(* IEC 61131-3 sources: SortJet_MasterSPS_Aufbau.fbsproj/07_Auftragsverwaltung/SystemCheck.prg.st^, 7 files *)

(* ---- Auftraege_Shuttle.meth.st ---- *)
(* METADATA
{
	"v3Meta": {
		"objectGuid": "9ff2d478-3fef-409c-b42e-3dce6a33e4ba"
	}
}
*)
METHOD PRIVATE Auftraege_Shuttle : BOOL
VAR_INPUT
  wpAutomatikkreis : WORD;
END_VAR

//-------------------------------------------------------------------------------------------------
// SYSTEMCHECK - AUTOMATIKKREIS 1
//-------------------------------------------------------------------------------------------------

Auftraege_Shuttle := FALSE;

FOR wlIndex := cERSTES_SHUTTLE TO cLETZTES_SHUTTLE DO
  IF wpAutomatikkreis = starrShuttleBasisParameter[wlIndex].stMKs.eaAutomatikkreis[1] THEN
    IF starrShuttleBasisParameter[wlIndex].stMKs.eStationsTyp = eInputshuttle THEN//101,102
      CASE starrShuttleBasisParameter[wlIndex].pAuftrag[cWAND_1].wTransferstationsNr1 OF

        cERSTE_STATION..cLETZTE_STATION:
          starrShuttleBasisParameter[wlIndex].pAuftrag[cWAND_1].stAuftragsOptionen.eGlastransport := eGlastransport_AufEinlaufVorab;
          starrShuttleBasisParameter[wlIndex].pAuftrag[cWAND_1].stAuftragsOptionen.eKippen_SollPosition := eKippen_Position_90Grad;
          Auftraege_Shuttle := TRUE;

        cERSTES_TRANSFERSHUTTLE..cLETZTES_TRANSFERSHUTTLE,
        cSPEICHER_1..cSPEICHER_2:
          starrShuttleBasisParameter[wlIndex].pAuftrag[cWAND_1].stAuftragsOptionen.eGlastransport := eGlastransport_AufAuslauf;
          starrShuttleBasisParameter[wlIndex].pAuftrag[cWAND_1].stAuftragsOptionen.eKippen_SollPosition := eKippen_Position_90Grad;//1.5
          Auftraege_Shuttle := TRUE;

        cERSTE_FAECHERWAGENSTATIONS_NR..cLETZTE_FAECHERWAGENSTATIONS_NR:
          starrShuttleBasisParameter[wlIndex].pAuftrag[cWAND_1].stAuftragsOptionen.eGlastransport := eGlastransport_AufAuslauf;
          starrShuttleBasisParameter[wlIndex].pAuftrag[cWAND_1].stAuftragsOptionen.eKippen_SollPosition := eKippen_Position_90Grad;
          Auftraege_Shuttle := TRUE;

        ELSE
          starrShuttleBasisParameter[wlIndex].pAuftrag[cWAND_1].stAuftragsOptionen.eGlastransport := eGlastransport_AufAuslauf;
          starrShuttleBasisParameter[wlIndex].pAuftrag[cWAND_1].stAuftragsOptionen.eKippen_SollPosition := eKippen_Position_90Grad;
          Auftraege_Shuttle := TRUE;

      END_CASE

    ELSIF starrShuttleBasisParameter[wlIndex].stMKs.eStationsTyp = eOutputshuttle THEN//103,104
      CASE starrShuttleBasisParameter[wlIndex].pAuftrag[cWAND_1].wTransferstationsNr1 OF

        cERSTES_TRANSFERSHUTTLE..cLETZTES_TRANSFERSHUTTLE,
        cSPEICHER_1:
          starrShuttleBasisParameter[wlIndex].pAuftrag[cWAND_1].stAuftragsOptionen.eGlastransport := eGlastransport_AufEinlaufVorab;
          starrShuttleBasisParameter[wlIndex].pAuftrag[cWAND_1].stAuftragsOptionen.eKippen_SollPosition := eKippen_Position_90Grad;//1.5
          Auftraege_Shuttle := TRUE;

        cERSTE_STATION..cLETZTE_STATION:
          starrShuttleBasisParameter[wlIndex].pAuftrag[cWAND_1].stAuftragsOptionen.eGlastransport := eGlastransport_AufAuslauf;
          starrShuttleBasisParameter[wlIndex].pAuftrag[cWAND_1].stAuftragsOptionen.eKippen_SollPosition := eKippen_Position_90Grad;
          Auftraege_Shuttle := TRUE;

        cERSTE_FAECHERWAGENSTATIONS_NR..cLETZTE_FAECHERWAGENSTATIONS_NR:
          starrShuttleBasisParameter[wlIndex].pAuftrag[cWAND_1].stAuftragsOptionen.eGlastransport := eGlastransport_AufAuslauf;
          starrShuttleBasisParameter[wlIndex].pAuftrag[cWAND_1].stAuftragsOptionen.eKippen_SollPosition := eKippen_Position_90Grad;
          Auftraege_Shuttle := TRUE;

        ELSE
          starrShuttleBasisParameter[wlIndex].pAuftrag[cWAND_1].stAuftragsOptionen.eGlastransport := eGlastransport_AufEinlaufVorab;
          starrShuttleBasisParameter[wlIndex].pAuftrag[cWAND_1].stAuftragsOptionen.eKippen_SollPosition := eKippen_Position_90Grad;
          Auftraege_Shuttle := TRUE;

      END_CASE
    ELSE
      starrShuttleBasisParameter[wlIndex].pAuftrag[cWAND_1].stAuftragsOptionen.eGlastransport := eGlastransport_AufEinlaufVorab;
      starrShuttleBasisParameter[wlIndex].pAuftrag[cWAND_1].stAuftragsOptionen.eKippen_SollPosition := eKippen_Default;
      Auftraege_Shuttle := TRUE;

    END_IF
  END_IF
END_FOR
END_METHOD

(* ---- Meldungen.act.st ---- *)
(* METADATA
{
	"v3Meta": {
		"objectGuid": "33333473-e459-491c-a043-28f329bb58b7"
	}
}
*)
ACTION Meldungen
//-------------------------------------------------------------------------------------------------
// MELDUNGEN
//-------------------------------------------------------------------------------------------------
(* Hinweis:
   - WatchIO
*)
FOR wlIndexAutomatikkreis := cERSTER_AUTOMATIKKREIS TO cLETZTER_AUTOMATIKKREIS DO
  WatchIo( (abpCheck[wlIndexAutomatikkreis] ) AND NOT M_Init_Ok, ioccCheckWaitInit);
  // -1 da die ioccKonstante bei AK 1 anfängt (Konstante AK1 = 1 ; somit würde die ioccKonstante + AK einen AK zu weit melden)
  WatchIo( ( abpCheck[wlIndexAutomatikkreis] ) AND NOT checkSafetyCircuitsClosedFromAutomaticCircuit(wlIndexAutomatikkreis, TRUE) AND NOT bgSicherheitstechnikBruecken, ( ioccCheckWaitSK_AK1 + wlIndexAutomatikkreis - 1) );
END_FOR

WatchIo( blCheckAktiv AND NOT M_Init_Ok, ioccCheckWaitInit);
END_ACTION

(* ---- Quittierung_Scheiben.act.st ---- *)
(* METADATA
{
	"v3Meta": {
		"objectGuid": "2a70e2fa-dcda-4b8f-820f-05f7864c9862"
	}
}
*)
ACTION Quittierung_Scheiben
//-------------------------------------------------------------------------------------------------
// QUITTIEREN DER SCHEIBEN IM SYSTEMCHECK [VERBUND]
//-------------------------------------------------------------------------------------------------

(* Hinweis:
   - Meldet eine Station im Systemcheck eine Scheibe [bQuittScheibe], wird sie wie im Auftrag quittiert
   - Die Richtung gibt das eigene Verbund- Flag der Station vor, der Partner steht in der Kopplung des Glasinterface
     [fest aus dem MK oder dynamisch aus Steuerung_VerbundCheck]
   - Check mit Vorgaenger: Die Station ist das Ziel, der Vorgaenger [aEintransporte] ist die Quelle
   - Check mit Nachfolger: Die Station ist die Quelle, der Nachfolger [aAustransporte] ist das Ziel
   - Quittiert wird nur, wenn die Station fuer den Partner quittiert [bStationQuittiertScheibe]
*)
FOR wlIndexQuitt := cERSTER_AUTOMATIKKREIS TO cLETZTER_AUTOMATIKKREIS DO

  IF ( abpCheck[wlIndexQuitt] ) THEN

    FOR wlIndexQuittStation := cERSTE_STATION TO cLETZTE_STATION DO

      stlQuittStation REF= getBasis( wlIndexQuittStation );

      IF    StationInAutomatikkreis( stlQuittStation.stMKs.eaAutomatikkreis, wlIndexQuitt )
            AND stlQuittStation.OutGlasTransport[cWAND_1].bQuittScheibe
      THEN

        // Eintransport: Station = Ziel
        IF stlQuittStation.bCheckMitVorgaenger[cWAND_1] THEN

          wlIndexQuittPartner := stlQuittStation.InGlasTransportVorgaenger[cWAND_1].stStationsNummern.NummerIntern;

          IF PruefungWertImIntervall( wlIndexQuittPartner, cERSTES_SHUTTLE, cLETZTE_FREMDANLAGE_EINLAUF ) THEN
            IF    ( stlQuittStation.stMKs.stSchnittstellendaten.aEintransporte.Station[wlIndexQuittPartner] <> TransportRichtung_EN.Default )
                  AND stlQuittStation.stMKs.stSchnittstellendaten.aEintransporte.bStationQuittiertScheibe[wlIndexQuittPartner]
            THEN
              ScheibenQuittierung( wpQuellstation := wlIndexQuittPartner,
                                   wpZielStation  := wlIndexQuittStation );
            END_IF
          END_IF

        // Austransport: Station = Quelle
        ELSIF stlQuittStation.bCheckMitNachfolger[cWAND_1] THEN

          wlIndexQuittPartner := stlQuittStation.InGlasTransportNachfolger[cWAND_1].stStationsNummern.NummerIntern;

          IF PruefungWertImIntervall( wlIndexQuittPartner, cERSTES_SHUTTLE, cLETZTE_FREMDANLAGE_EINLAUF ) THEN
            IF    ( stlQuittStation.stMKs.stSchnittstellendaten.aAustransporte.Station[wlIndexQuittPartner] <> TransportRichtung_EN.Default )
                  AND stlQuittStation.stMKs.stSchnittstellendaten.aAustransporte.bStationQuittiertScheibe[wlIndexQuittPartner]
            THEN
              IF stlQuittStation.stMKs.stSchnittstellendaten.bStationIstShuttle THEN
                ScheibenQuittierung( wpQuellstation := wlIndexQuittStation,
                                     wpZielStation  := wlIndexQuittPartner,
                                     wpAuftragsTyp  := 1 );
              ELSE
                ScheibenQuittierung( wpQuellstation := wlIndexQuittStation,
                                     wpZielStation  := wlIndexQuittPartner );
              END_IF
            END_IF
          END_IF

        END_IF

      END_IF

    END_FOR

  END_IF

END_FOR
END_ACTION

(* ---- Reset.act.st ---- *)
(* METADATA
{
	"v3Meta": {
		"objectGuid": "c82983ad-c0e7-4e08-a2e4-b90c50d3f8d7"
	}
}
*)
ACTION Reset
//-------------------------------------------------------------------------------------------------
// RESET
//-------------------------------------------------------------------------------------------------
(* Hinweis:
   - Fehlerbit zuruecksetzen
   - Shuttledatenbit zuruecksetzen
   - Merker zuruecksetzen [Welches Transfershuttle benutzt wurde]
*)
FOR wlIndexAutomatikkreis := cERSTER_AUTOMATIKKREIS TO cLETZTER_AUTOMATIKKREIS DO

  IF ( abpReset[wlIndexAutomatikkreis] ) THEN

    abpFehler[wlIndexAutomatikkreis] := FALSE;

    FOR wlIndexStationsnummer := cERSTES_SHUTTLE TO cLETZTES_SHUTTLE DO
      IF StationInAutomatikkreis(starrShuttleBasisParameter[wlIndexStationsnummer].stMKs.eaAutomatikkreis, wlIndexAutomatikkreis) THEN
        abpStationsDatenErhalten[wlIndexStationsnummer, cWAND_1] := FALSE;
        ablShuttleCheckAktiv[wlIndexStationsnummer] := FALSE;
      END_IF
    END_FOR

    FOR wlIndexStationsnummer := cERSTE_STATION TO cLETZTE_STATION DO
      IF StationInAutomatikkreis(starrStationBasisParameter[wlIndexStationsnummer].stMKs.eaAutomatikkreis, wlIndexAutomatikkreis) THEN
        abpStationsDatenErhalten[wlIndexStationsnummer, cWAND_1] := FALSE;
        ablStationCheckAktiv[wlIndexStationsnummer] := FALSE;
      END_IF
    END_FOR

    abpReset[wlIndexAutomatikkreis] := FALSE;

    wlAktiverZyklus := 1;

    FOR wlIndexSystemcheckZyklus := 1 TO wgAnzahlSystemcheckZyklen DO
      ablCheck[wlIndexAutomatikkreis, wlIndexSystemcheckZyklus] := FALSE;
      ablCheckDone[wlIndexAutomatikkreis, wlIndexSystemcheckZyklus] := FALSE;
    END_FOR

  END_IF

END_FOR
END_ACTION

(* ---- Steuerung_VerbundCheck.meth.st ---- *)
(* METADATA
{
	"v3Meta": {
		"objectGuid": "2106329f-ce22-4754-a4e1-a7a15d593805"
	}
}
*)
METHOD PRIVATE Steuerung_VerbundCheck : BOOL
VAR_INPUT
  wpAutomatikkreis : WORD;
  wpZyklus         : WORD;
END_VAR
VAR
  ilNachfolger        : INT;
  wlNachfolger        : WORD;
  wlVorgaenger        : WORD;
  wlPartner           : WORD;
  wlIndexAK           : WORD;
  wlIndexWand         : WORD;
  blVorgaengerImAK    : BOOL;
  blNachfolgerImAK    : BOOL;
  blPartnerPrueftMit  : BOOL;
  stlFesterPartner    : REFERENCE TO StationBasisParameter_ST;
END_VAR

(* Hinweis:
   - Liegt eine Scheibe ueber der Grenze zweier Stationen, pruefen beide Stationen gemeinsam
   - Ein Paar [Vorgaenger => Nachfolger] ergibt sich aus dem Eintransport des Nachfolgers [aEintransporte]
     und gilt, wenn der Auslaufsensor des Vorgaengers und der Einlaufsensor des Nachfolgers belegt sind
   - Ist der Vorgaenger eine Anlegestation [MK bIstAnlegestation], muss er genau eine Scheibe haben
   - Ein Nachfolger der schon mit seinem eigenen Nachfolger prueft, wird nicht zusaetzlich mit seinem Vorgaenger
     verbunden; deshalb wird von der letzten Station zur ersten Station gearbeitet [das Ende der Kette gewinnt]
   - Die Partner koennen in verschiedenen Automatikkreisen liegen; jeder Automatikkreis setzt nur die Flags
     seiner eigenen Stationen
   - Prueft der Automatikkreis des Partners nicht mit, muss er zusaetzlich den Systemcheck machen [Hinweis]
   - Hat eine Station im MK keinen festen Vorgaenger/Nachfolger [dynamisch oder default], wird die Kopplung
     des Glasinterface hier auf den Partner des Paars gesetzt [Job_Stationen koppelt nur feste Partner]
     Die Quittierung im Systemcheck leitet den Partner aus dieser Kopplung ab
*)
FOR ilNachfolger := WORD_TO_INT( cLETZTE_STATION ) TO WORD_TO_INT( cERSTE_STATION ) BY -1 DO

  wlNachfolger := INT_TO_WORD( ilNachfolger );

  FOR wlVorgaenger := cERSTE_STATION TO cLETZTE_STATION DO

    blVorgaengerImAK := StationInAutomatikkreis( starrStationBasisParameter[wlVorgaenger].stMKs.eaAutomatikkreis, wpAutomatikkreis );
    blNachfolgerImAK := StationInAutomatikkreis( starrStationBasisParameter[wlNachfolger].stMKs.eaAutomatikkreis, wpAutomatikkreis );

    IF    ( blVorgaengerImAK OR blNachfolgerImAK )
          AND ( wlVorgaenger <> wlNachfolger )
          AND ( starrStationBasisParameter[wlNachfolger].stMKs.stSchnittstellendaten.aEintransporte.Station[wlVorgaenger] <> TransportRichtung_EN.Default )
          AND starrStationBasisParameter[wlVorgaenger].OutGlasTransport[cWAND_1].bAuslaufsensor
          AND starrStationBasisParameter[wlNachfolger].OutGlasTransport[cWAND_1].bEinlaufsensor
          AND (    NOT starrStationBasisParameter[wlVorgaenger].stMKs.stStationsOptionen.stAnlegetisch.bIstAnlegestation
                OR ( starrStationBasisParameter[wlVorgaenger].pAuftrag[cWAND_1].wAnzahlScheiben = 1 ) )
          AND NOT starrStationBasisParameter[wlNachfolger].bCheckMitNachfolger[cWAND_1]
    THEN

      IF blVorgaengerImAK THEN
        starrStationBasisParameter[wlVorgaenger].bCheckMitNachfolger[cWAND_1] := TRUE;
      END_IF

      IF blNachfolgerImAK THEN
        starrStationBasisParameter[wlNachfolger].bCheckMitVorgaenger[cWAND_1] := TRUE;
      END_IF

      // Kopplung Glasinterface: Vorgaenger => Nachfolger
      stlFesterPartner REF= getBasis( starrStationBasisParameter[wlVorgaenger].stMKs.stSchnittstellendaten.wNachfolgerStation );
      IF NOT __ISVALIDREF( stlFesterPartner ) THEN
        FOR wlIndexWand := cWAND_1 TO cANZAHL_WAENDE DO
          starrStationBasisParameter[wlVorgaenger].InGlasTransportNachfolger[wlIndexWand] := starrStationBasisParameter[wlNachfolger].OutGlasTransport[cWAND_1];
        END_FOR
      END_IF

      // Kopplung Glasinterface: Nachfolger => Vorgaenger
      stlFesterPartner REF= getBasis( starrStationBasisParameter[wlNachfolger].stMKs.stSchnittstellendaten.wVorgaengerStation );
      IF NOT __ISVALIDREF( stlFesterPartner ) THEN
        FOR wlIndexWand := cWAND_1 TO cANZAHL_WAENDE DO
          starrStationBasisParameter[wlNachfolger].InGlasTransportVorgaenger[wlIndexWand] := starrStationBasisParameter[wlVorgaenger].OutGlasTransport[cWAND_1];
        END_FOR
      END_IF

      // Liegt nur eine der beiden Stationen im geprueften Automatikkreis, liegt der Partner in einem anderen
      // Automatikkreis und dieser muss den Systemcheck zusaetzlich machen
      IF NOT blVorgaengerImAK OR NOT blNachfolgerImAK THEN

        IF blVorgaengerImAK THEN
          wlPartner := wlNachfolger;
        ELSE
          wlPartner := wlVorgaenger;
        END_IF

        blPartnerPrueftMit := FALSE;
        FOR wlIndexAK := cERSTER_AUTOMATIKKREIS TO cANZAHL_AUTOMATIKKREISE DO
          IF starrStationBasisParameter[wlPartner].stMKs.eaAutomatikkreis[wlIndexAK] <> 0 THEN
            IF abpCheck[starrStationBasisParameter[wlPartner].stMKs.eaAutomatikkreis[wlIndexAK]] THEN
              blPartnerPrueftMit := TRUE;
            END_IF
          END_IF
        END_FOR

        IF NOT blPartnerPrueftMit THEN
          wpgFehlerdaten[0] := AutomatikkreisBestimmen( wlPartner );
          SpsHinweis( eFehler_Station,
                      cMELDUNG_SYSTEMCHECK_VERBUND_ANDERER_AK_NOETIG,
                      wlPartner,
                      wpAutomatikkreis,
                      wpgFehlerdaten );
        END_IF

      END_IF

    END_IF

  END_FOR

END_FOR

Steuerung_VerbundCheck := TRUE;
END_METHOD

(* ---- Systemcheck.meth.st ---- *)
(* METADATA
{
	"v3Meta": {
		"objectGuid": "db7a5787-dcad-4426-bbf6-73751d4de64b"
	}
}
*)
METHOD PRIVATE Systemcheck : BOOL
VAR_INPUT
  wpAutomatikkreis : WORD;
  wpZyklus         : WORD;
END_VAR

VAR

  blSystemcheckdatenErhalten : BOOL;

  wlIndex            : WORD;
  wlSubIndex         : WORD;
  wlIndexStationen   : WORD;
  wlStationOhneDaten : WORD; // Externe Stationsnummer der ersten Station ohne Auftragsdaten

END_VAR

//-------------------------------------------------------------------------------------------------
// SYSTEMCHECK - AUTOMATIKKREIS X
//-------------------------------------------------------------------------------------------------

IF ablCheck[wpAutomatikkreis, wpZyklus] THEN

  CASE asteplCheck[wpAutomatikkreis, wpZyklus] OF

    // SYSTEMCHECK ==================================
    STEP_0_E:
      (* Anmerkung:
         - -
      *)
      atonlWarnungSystemCheckBeginnt[wpAutomatikkreis](IN:= FALSE);
      atonlCheck[wpAutomatikkreis](IN := FALSE);

      IF ( NOT agbResetAktiv[wpAutomatikkreis] )THEN
        ailAnzahlShuttleCheckAktiv[wpAutomatikkreis]      := 0;
        ailAnzahlStationenCheckAktiv[wpAutomatikkreis]    := 0;
        ailAnzahlFWStationenCheckAktiv[wpAutomatikkreis]  := 0;

        ablTimeOutMeldungGenerieren[wpAutomatikkreis] := TRUE;
        ablStationFehlerImCheck[wpAutomatikkreis]     := FALSE;

        // Status zurueck setzen
        FOR wlIndex := cERSTE_STATION TO cLETZTE_STATION DO
          IF    ( StationInAutomatikkreis(starrStationBasisParameter[wlIndex].stMKs.eaAutomatikkreis, wpAutomatikkreis) )
                AND ( starrStationBasisParameter[wlIndex].stMKs.eSystemcheckZyklus = wpZyklus )
          THEN
            ablStationCheckAktiv[wlIndex] := FALSE;
          END_IF
        END_FOR

        FOR wlIndex := cERSTES_SHUTTLE TO cLETZTES_SHUTTLE DO
          IF    ( StationInAutomatikkreis(starrShuttleBasisParameter[wlIndex].stMKs.eaAutomatikkreis, wpAutomatikkreis) )
                AND ( starrShuttleBasisParameter[wlIndex].stMKs.eSystemcheckZyklus = wpZyklus )
          THEN
            ablShuttleCheckAktiv[wlIndex] := FALSE;
          END_IF
        END_FOR

        FOR wlIndex := cERSTE_FAECHERWAGENSTATIONS_NR TO cLETZTE_FAECHERWAGENSTATIONS_NR DO
          IF    ( StationInAutomatikkreis(starrFaecherwagenBasisParameter[wlIndex].stMKs.eaAutomatikkreis, wpAutomatikkreis) )
                AND ( starrFaecherwagenBasisParameter[wlIndex].stMKs.eSystemcheckZyklus = wpZyklus )
          THEN
            ablFWCheckAktiv[wlIndex] := FALSE;
          END_IF
        END_FOR

        IF NOT TransferShuttleBetriebsstopAktiv(wpAutomatikkreis) THEN
          asteplCheck[wpAutomatikkreis, wpZyklus] := STEP_10_E;
        ELSE
          SpsError( eFehler_Station,
                    cMELDUNG_SYSTEMCHECK_NICHT_MOEGLICH_TS_BETRIEBSSTOP,
                    0,
                    wpAutomatikkreis,
                    wpgFehlerdaten );
          asteplCheck[wpAutomatikkreis, wpZyklus] := STEP_900_E;
        END_IF
      END_IF

    // SYSTEMCHECK ==================================
    STEP_10_E:
      (* Hinweis:
         - SystemCheck starten sobald;
           => Daten eingetroffen sind
           => Sicherheitskreise / Druckluft / NotAus etc. okay melden
      *)
      IF (  atonlWaitCheck[wpAutomatikkreis].Q  ) THEN
        atonlCheckWarteAufMMIDaten[wpAutomatikkreis]( IN :=  FALSE );
        asteplCheck[wpAutomatikkreis, wpZyklus] := STEP_20_E;
      END_IF

    // SYSTEMCHECK ==================================
    STEP_20_E:
      (* Hinweis:
         - SystemCheck starten sobald;
           => Daten eingetroffen sind
           => Sicherheitskreise / Druckluft / NotAus etc. okay melden
      *)
      blSystemcheckdatenErhalten := TRUE;
      wlStationOhneDaten := 0;

      FOR wlIndexStationen := cERSTE_STATION TO cLETZTE_STATION DO
        IF ( starrStationBasisParameter[wlIndexStationen].stMKs.eSystemcheckZyklus = wpZyklus )
           AND ( StationInAutomatikkreis(starrStationBasisParameter[wlIndexStationen].stMKs.eaAutomatikkreis, wpAutomatikkreis) )
           AND ( NOT starrStationBasisParameter[wlIndexStationen].stMKs.bDeaktivieren )
        THEN
          IF NOT abpStationsDatenErhalten[wlIndexStationen, cWAND_1] THEN
            blSystemcheckdatenErhalten := FALSE;
            IF ( wlStationOhneDaten = 0 ) THEN
              wlStationOhneDaten := starrStationBasisParameter[wlIndexStationen].stMKs.stStationsNummern.NummerExtern;
            END_IF
          END_IF
        END_IF
      END_FOR

      FOR wlIndexStationen := cERSTES_SHUTTLE TO cLETZTES_SHUTTLE DO
        IF (starrShuttleBasisParameter[wlIndexStationen].stMKs.eSystemcheckZyklus = wpZyklus )
           AND ( StationInAutomatikkreis(starrShuttleBasisParameter[wlIndexStationen].stMKs.eaAutomatikkreis, wpAutomatikkreis) )
           AND ( NOT starrShuttleBasisParameter[wlIndexStationen].stMKs.bDeaktivieren )
        THEN
          IF NOT abpStationsDatenErhalten[wlIndexStationen, cWAND_1] THEN
            blSystemcheckdatenErhalten := FALSE;
            IF ( wlStationOhneDaten = 0 ) THEN
              wlStationOhneDaten := starrShuttleBasisParameter[wlIndexStationen].stMKs.stStationsNummern.NummerExtern;
            END_IF
          END_IF
        END_IF
      END_FOR

      IF blSystemcheckdatenErhalten OR bgInbetriebnahmeBit THEN
        atonlCheckWarteAufMMIDaten[wpAutomatikkreis]( IN :=  FALSE );
        asteplCheck[wpAutomatikkreis, wpZyklus] := STEP_30_E;
      END_IF

      (* Hinweis:
         - Nicht alle Daten in der vorgeschriebenen Zeit eingetroffen
      *)
      atonlCheckWarteAufMMIDaten[wpAutomatikkreis]( IN :=  TRUE, PT := T#5S);
      IF atonlCheckWarteAufMMIDaten[wpAutomatikkreis].Q THEN
        atonlCheckWarteAufMMIDaten[wpAutomatikkreis]( IN :=  FALSE );
        wpgFehlerdaten[0] := wlStationOhneDaten;
        SpsError( eFehler_Station,
                  cMELDUNG_SYSTEMCHECK_AUFTRAGSDATEN_TIMEOUT,
                  0,
                  wpAutomatikkreis,
                  wpgFehlerdaten );

        asteplCheck[wpAutomatikkreis, wpZyklus] := STEP_900_E;
      END_IF

    // SYSTEMCHECK ==================================
    STEP_30_E:
      (* Hinweis:
         - Vor dem Starten des SystemChecks wird ein akustisches Signal ausgegeben [Horn]
           => 3 - 5 Sekunden zur Fluchtmoeglichkeit geben bevor die Anlage gestartet wird [Fals noch jemand im Sicherheitskreis ist]
      *)
      FOR wlSubIndex := 1 TO cANZAHL_HUPEN DO
        Horn_AK[wpAutomatikkreis,wlSubIndex].wpStatusArt      := 1;
        Horn_AK[wpAutomatikkreis,wlSubIndex].tpHornZeit       := T#3S;
        Horn_AK[wpAutomatikkreis,wlSubIndex].bpHornAktivieren := TRUE;
      END_FOR

      atonlWarnungSystemCheckBeginnt[wpAutomatikkreis]( IN := TRUE,
                                                        PT := T#3s );

      IF ( atonlWarnungSystemCheckBeginnt[wpAutomatikkreis].Q ) THEN
        atonlWarnungSystemCheckBeginnt[wpAutomatikkreis](IN:= FALSE);
        asteplCheck[wpAutomatikkreis, wpZyklus] := STEP_40_E;
      END_IF

    // SYSTEMCHECK ==================================
    STEP_40_E:
      (* Hinweis:
         - Verbund- SystemCheck
      *)
      Steuerung_VerbundCheck( wpAutomatikkreis, wpZyklus );

      (* Hinweis:
         - Zuweisen der Systemcheckdaten
      *)
      FOR wlIndexStationen := cERSTE_STATION TO cLETZTE_STATION DO
        IF    starrStationBasisParameter[wlIndexStationen].stMKs.eSystemcheckZyklus = wpZyklus
              AND StationInAutomatikkreis(starrStationBasisParameter[wlIndexStationen].stMKs.eaAutomatikkreis, wpAutomatikkreis)
        THEN
          starrStationBasisParameter[wlIndexStationen].pAuftrag[cWAND_1] := abgDateStationCheck[wlIndexStationen, cWAND_1];
        END_IF
      END_FOR

      FOR wlIndexStationen := cERSTES_SHUTTLE TO cLETZTES_SHUTTLE DO
        IF    starrShuttleBasisParameter[wlIndexStationen].stMKs.eSystemcheckZyklus = wpZyklus
              AND StationInAutomatikkreis(starrShuttleBasisParameter[wlIndexStationen].stMKs.eaAutomatikkreis, wpAutomatikkreis)
        THEN
          starrShuttleBasisParameter[wlIndexStationen].pAuftrag[cWAND_1] := abgDateStationCheck[wlIndexStationen, cWAND_1];
        END_IF
      END_FOR

      // Auftragsdaten aufbereiten
      Auftraege_Shuttle( wpAutomatikkreis );

      (* Hinweis:
         - Starten des Baustein- SystemChecks
      *)
      // STATION
      FOR wlIndex := cERSTE_STATION TO cLETZTE_STATION DO

        IF   StationInAutomatikkreis(starrStationBasisParameter[wlIndex].stMKs.eaAutomatikkreis, wpAutomatikkreis)
             AND (   starrStationBasisParameter[wlIndex].stMKs.eSystemcheckZyklus = wpZyklus
                   OR starrStationBasisParameter[wlIndex].bCheckMitVorgaenger[cWAND_1]
                   OR starrStationBasisParameter[wlIndex].bCheckMitNachfolger[cWAND_1] )
        THEN
          starrStationBasisParameter[wlIndex].bCheck := TRUE;
          ailAnzahlStationenCheckAktiv[wpAutomatikkreis] := ailAnzahlStationenCheckAktiv[wpAutomatikkreis] + 1;
          ablStationCheckAktiv[wlIndex] := TRUE;
        END_IF

      END_FOR

      // SHUTTLE
      FOR wlIndex := cERSTES_SHUTTLE TO cLETZTES_SHUTTLE DO

        IF StationInAutomatikkreis(starrShuttleBasisParameter[wlIndex].stMKs.eaAutomatikkreis, wpAutomatikkreis)
           AND (   starrShuttleBasisParameter[wlIndex].stMKs.eSystemcheckZyklus = wpZyklus
                 OR starrShuttleBasisParameter[wlIndex].bCheckMitVorgaenger[cWAND_1]
                 OR starrShuttleBasisParameter[wlIndex].bCheckMitNachfolger[cWAND_1] )
        THEN
          starrShuttleBasisParameter[wlIndex].bCheck := TRUE;
          ailAnzahlShuttleCheckAktiv[wpAutomatikkreis] := ailAnzahlShuttleCheckAktiv[wpAutomatikkreis] + 1;
          ablShuttleCheckAktiv[wlIndex] := TRUE;
        END_IF

      END_FOR

      // FW
      FOR wlIndex := cERSTE_FAECHERWAGENSTATIONS_NR TO cLETZTE_FAECHERWAGENSTATIONS_NR DO

        IF StationInAutomatikkreis(starrFaecherwagenBasisParameter[wlIndex].stMKs.eaAutomatikkreis, wpAutomatikkreis)
           AND ( starrFaecherwagenBasisParameter[wlIndex].stMKs.eSystemcheckZyklus = wpZyklus  )
        THEN
          starrFaecherwagenBasisParameter[wlIndex].bCheck := TRUE;
          ailAnzahlFWStationenCheckAktiv[wpAutomatikkreis] := ailAnzahlFWStationenCheckAktiv[wpAutomatikkreis] + 1;
          ablFWCheckAktiv[wlIndex] := TRUE;
        END_IF

      END_FOR

      asteplCheck[wpAutomatikkreis, wpZyklus] := STEP_100_E;

    // SYSTEMCHECK ==================================
    STEP_100_E:
      (* Hinweis:
         - Initalisierung des Timers fuer dei SystemCheck Ueberwachung
      *)
      atonlCheck[wpAutomatikkreis](IN := TRUE, PT := tgTimeWarteAufCheckDone );

      (* Hinweis:
         - Warten bis die Stationen [Einlaufstrecke] ihren SystemCheck beendet haben
      *)
      // SHUTTLE
      FOR wlIndex := cERSTES_SHUTTLE TO cLETZTES_SHUTTLE DO

        IF StationInAutomatikkreis(starrShuttleBasisParameter[wlIndex].stMKs.eaAutomatikkreis, wpAutomatikkreis)
           AND (   starrShuttleBasisParameter[wlIndex].stMKs.eSystemcheckZyklus = wpZyklus
                 OR starrShuttleBasisParameter[wlIndex].bCheckMitVorgaenger[cWAND_1]
                 OR starrShuttleBasisParameter[wlIndex].bCheckMitNachfolger[cWAND_1] )
        THEN

          IF (   starrShuttleBasisParameter[wlIndex].bCheckAbgeschlossen
               AND starrShuttleBasisParameter[wlIndex].bCheck )
          THEN
            starrShuttleBasisParameter[wlIndex].bCheck := FALSE;
            ailAnzahlShuttleCheckAktiv[wpAutomatikkreis] := ailAnzahlShuttleCheckAktiv[wpAutomatikkreis] - 1;
            ablShuttleCheckAktiv[wlIndex] := FALSE;
          END_IF

        END_IF

      END_FOR

      // STATION
      FOR wlIndex :=   cERSTE_STATION TO cLETZTE_STATION DO

        IF StationInAutomatikkreis(starrStationBasisParameter[wlIndex].stMKs.eaAutomatikkreis, wpAutomatikkreis)
           AND (   starrStationBasisParameter[wlIndex].stMKs.eSystemcheckZyklus = wpZyklus
                 OR starrStationBasisParameter[wlIndex].bCheckMitVorgaenger[cWAND_1]
                 OR starrStationBasisParameter[wlIndex].bCheckMitNachfolger[cWAND_1] )
        THEN

          IF (   starrStationBasisParameter[wlIndex].bCheckAbgeschlossen
               AND starrStationBasisParameter[wlIndex].bCheck )
          THEN
            starrStationBasisParameter[wlIndex].bCheck := FALSE;
            ailAnzahlStationenCheckAktiv[wpAutomatikkreis] := ailAnzahlStationenCheckAktiv[wpAutomatikkreis] - 1;
            ablStationCheckAktiv[wlIndex] := FALSE;
          END_IF

        END_IF

      END_FOR

      // FW
      FOR wlIndex := cERSTE_FAECHERWAGENSTATIONS_NR TO cLETZTE_FAECHERWAGENSTATIONS_NR DO

        IF StationInAutomatikkreis(starrFaecherwagenBasisParameter[wlIndex].stMKs.eaAutomatikkreis, wpAutomatikkreis)
           AND (   starrFaecherwagenBasisParameter[wlIndex].stMKs.eSystemcheckZyklus = wpZyklus  )
        THEN

          IF (   starrFaecherwagenBasisParameter[wlIndex].bCheckAbgeschlossen
               AND starrFaecherwagenBasisParameter[wlIndex].bCheck )
          THEN
            starrFaecherwagenBasisParameter[wlIndex].bCheck := FALSE;
            ailAnzahlFWStationenCheckAktiv[wpAutomatikkreis] := ailAnzahlFWStationenCheckAktiv[wpAutomatikkreis] - 1;
            ablFWCheckAktiv[wlIndex] := FALSE;
          END_IF

        END_IF

      END_FOR

      IF (  ailAnzahlShuttleCheckAktiv[wpAutomatikkreis]         = 0
           AND ailAnzahlStationenCheckAktiv[wpAutomatikkreis]       = 0
           AND ailAnzahlFWStationenCheckAktiv[wpAutomatikkreis]     = 0 )
      THEN
        (* Hinweis:
           - Alle Stationen haben den Check beendet, Stationen mit Fehler wurden bereits gemeldet
        *)
        IF ( ablStationFehlerImCheck[wpAutomatikkreis] ) THEN
          asteplCheck[wpAutomatikkreis, wpZyklus] := STEP_900_E;
        ELSE
          asteplCheck[wpAutomatikkreis, wpZyklus] := STEP_1000_E;
        END_IF

      END_IF

      // zeitliche Überwachung des Systemchecks !
      IF ( atonlCheck[wpAutomatikkreis].Q ) THEN

        // SHUTTLE
        FOR wlIndex := cERSTES_SHUTTLE TO cLETZTES_SHUTTLE DO

          IF StationInAutomatikkreis(starrShuttleBasisParameter[wlIndex].stMKs.eaAutomatikkreis, wpAutomatikkreis)
             AND starrShuttleBasisParameter[wlIndex].bCheck
          THEN
            starrShuttleBasisParameter[wlIndex].bCheck := FALSE;

            IF ( NOT starrShuttleBasisParameter[wlIndex].bCheckAbgeschlossen ) THEN
              ablTimeOutMeldungGenerieren[wpAutomatikkreis] := FALSE;
              wpgFehlerdaten[0] := wlIndex;
              SpsError( eFehler_Station,
                        cMELDUNG_SYSTEMCHECK_STATION_BEENDET_DIESEN_NICHT,
                        wlIndex,
                        AutomatikkreisBestimmen(wlIndex),
                        starrShuttleBasisParameter[wlIndex].awFehlerInformationen );
            END_IF

          END_IF

        END_FOR

        // STATION
        FOR wlIndex :=   cERSTE_STATION TO cLETZTE_STATION DO

          IF StationInAutomatikkreis(starrStationBasisParameter[wlIndex].stMKs.eaAutomatikkreis, wpAutomatikkreis)
             AND starrStationBasisParameter[wlIndex].bCheck
          THEN
            starrStationBasisParameter[wlIndex].bCheck := FALSE;

            IF ( NOT starrStationBasisParameter[wlIndex].bCheckAbgeschlossen ) THEN
              ablTimeOutMeldungGenerieren[wpAutomatikkreis] := FALSE;
              wpgFehlerdaten[0] := wlIndex;
              SpsError( eFehler_Station,
                        cMELDUNG_SYSTEMCHECK_STATION_BEENDET_DIESEN_NICHT,
                        wlIndex,
                        AutomatikkreisBestimmen(wlIndex),
                        starrStationBasisParameter[wlIndex].awFehlerInformationen );
            END_IF

          END_IF

        END_FOR

        // FW
        FOR wlIndex := cERSTE_FAECHERWAGENSTATIONS_NR TO cLETZTE_FAECHERWAGENSTATIONS_NR DO

          IF StationInAutomatikkreis(starrFaecherwagenBasisParameter[wlIndex].stMKs.eaAutomatikkreis, wpAutomatikkreis)
             AND starrFaecherwagenBasisParameter[wlIndex].bCheck
          THEN
            starrFaecherwagenBasisParameter[wlIndex].bCheck := FALSE;

            IF ( NOT starrFaecherwagenBasisParameter[wlIndex].bCheckAbgeschlossen ) THEN
              ablTimeOutMeldungGenerieren[wpAutomatikkreis] := FALSE;
              wpgFehlerdaten[0] := wlIndex;
              SpsError( eFehler_Station,
                        cMELDUNG_SYSTEMCHECK_STATION_BEENDET_DIESEN_NICHT,
                        wlIndex,
                        AutomatikkreisBestimmen(wlIndex),
                        starrFaecherwagenBasisParameter[wlIndex].awFehlerInformationen );
            END_IF

          END_IF

        END_FOR

        (* Hinweis:
           - Time Out Fehler generieren wenn sonst kein Fehler generiert wurde
        *)
        IF ( ablTimeOutMeldungGenerieren[wpAutomatikkreis] ) THEN
          wpgFehlerdaten[0] := wpAutomatikkreis;
          SpsHinweis( eFehler_Station,
                      cMELDUNG_SYSTEMCHECK_TIMEOUT,
                      0,
                      AutomatikkreisBestimmen(wpAutomatikkreis),
                      wpgFehlerdaten );
        END_IF

        asteplCheck[wpAutomatikkreis, wpZyklus] := STEP_900_E;

      END_IF

      // Fehler:
      //   - Bausteinfehler waerend des SystemCheks
      // SHUTTLE
      FOR wlIndex := cERSTES_SHUTTLE TO cLETZTES_SHUTTLE DO

        IF StationInAutomatikkreis(starrShuttleBasisParameter[wlIndex].stMKs.eaAutomatikkreis, wpAutomatikkreis)
           AND starrShuttleBasisParameter[wlIndex].bFehler
           AND starrShuttleBasisParameter[wlIndex].bCheck
        THEN
          starrShuttleBasisParameter[wlIndex].bCheck := FALSE;
          wpgFehlerdaten[0] := starrShuttleBasisParameter[wlIndex].wFehlerNummer;
          SpsError( eFehler_Station,
                    starrShuttleBasisParameter[wlIndex].wFehlerNummer,
                    wlIndex,
                    AutomatikkreisBestimmen(wlIndex),
                    starrShuttleBasisParameter[wlIndex].awFehlerInformationen );

          ailAnzahlShuttleCheckAktiv[wpAutomatikkreis] := ailAnzahlShuttleCheckAktiv[wpAutomatikkreis] - 1;
          ablShuttleCheckAktiv[wlIndex]                := FALSE;
          ablStationFehlerImCheck[wpAutomatikkreis]    := TRUE;

        END_IF

      END_FOR

      // STATION
      FOR wlIndex :=   cERSTE_STATION TO cLETZTE_STATION DO

        IF StationInAutomatikkreis(starrStationBasisParameter[wlIndex].stMKs.eaAutomatikkreis, wpAutomatikkreis)
           AND starrStationBasisParameter[wlIndex].bFehler
           AND starrStationBasisParameter[wlIndex].bCheck
        THEN
          starrStationBasisParameter[wlIndex].bCheck := FALSE;
          wpgFehlerdaten[0] := starrStationBasisParameter[wlIndex].wFehlerNummer;
          SpsError( eFehler_Station,
                    starrStationBasisParameter[wlIndex].wFehlerNummer,
                    wlIndex,
                    AutomatikkreisBestimmen(wlIndex),
                    starrStationBasisParameter[wlIndex].awFehlerInformationen );

          ailAnzahlStationenCheckAktiv[wpAutomatikkreis] := ailAnzahlStationenCheckAktiv[wpAutomatikkreis] - 1;
          ablStationCheckAktiv[wlIndex]                  := FALSE;
          ablStationFehlerImCheck[wpAutomatikkreis]      := TRUE;
        END_IF

      END_FOR

      // FW
      FOR wlIndex :=   cERSTE_FAECHERWAGENSTATIONS_NR TO cLETZTE_FAECHERWAGENSTATIONS_NR DO

        IF StationInAutomatikkreis(starrFaecherwagenBasisParameter[wlIndex].stMKs.eaAutomatikkreis, wpAutomatikkreis)
           AND starrFaecherwagenBasisParameter[wlIndex].bFehler
           AND starrFaecherwagenBasisParameter[wlIndex].bCheck
        THEN
          starrFaecherwagenBasisParameter[wlIndex].bCheck := FALSE;
          wpgFehlerdaten[0] := starrFaecherwagenBasisParameter[wlIndex].wFehlerNummer;
          SpsError( eFehler_Station,
                    starrFaecherwagenBasisParameter[wlIndex].wFehlerNummer,
                    wlIndex,
                    AutomatikkreisBestimmen(wlIndex),
                    starrFaecherwagenBasisParameter[wlIndex].awFehlerInformationen );

          ailAnzahlFWStationenCheckAktiv[wpAutomatikkreis] := ailAnzahlFWStationenCheckAktiv[wpAutomatikkreis] - 1;
          ablFWCheckAktiv[wlIndex]                         := FALSE;
          ablStationFehlerImCheck[wpAutomatikkreis]        := TRUE;
        END_IF

      END_FOR

    // SYSTEMCHECK ==================================
    STEP_900_E:
      abpFehler[wpAutomatikkreis] := TRUE;
      ablCheck[wpAutomatikkreis, wpZyklus] := FALSE;

    // SYSTEMCHECK ==================================
    STEP_1000_E:
      abpFehler[wpAutomatikkreis] := FALSE;
      ablCheckDone[wpAutomatikkreis, wpZyklus] := TRUE;

  // SYSTEMCHECK ==================================
  END_CASE

ELSIF ( asteplCheck[wpAutomatikkreis, wpZyklus] <> STEP_0_E ) THEN

  ablCheckDone[wpAutomatikkreis, wpZyklus] := FALSE;

  // SHUTTLE
  FOR wlIndex := cERSTES_SHUTTLE TO cLETZTES_SHUTTLE DO
    IF StationInAutomatikkreis(starrShuttleBasisParameter[wlIndex].stMKs.eaAutomatikkreis, wpAutomatikkreis) THEN
      starrShuttleBasisParameter[wlIndex].bCheck := FALSE;
    END_IF
  END_FOR

  // STATION
  FOR wlIndex :=   cERSTE_STATION TO cLETZTE_STATION DO
    IF StationInAutomatikkreis(starrStationBasisParameter[wlIndex].stMKs.eaAutomatikkreis, wpAutomatikkreis) THEN
      starrStationBasisParameter[wlIndex].bCheck := FALSE;
    END_IF
  END_FOR

  // FW
  FOR wlIndex :=   cERSTE_FAECHERWAGENSTATIONS_NR TO cLETZTE_FAECHERWAGENSTATIONS_NR DO
    IF StationInAutomatikkreis(starrFaecherwagenBasisParameter[wlIndex].stMKs.eaAutomatikkreis, wpAutomatikkreis) THEN
      starrFaecherwagenBasisParameter[wlIndex].bCheck := FALSE;
    END_IF
  END_FOR

  ailAnzahlShuttleCheckAktiv[wpAutomatikkreis]      := 0;
  ailAnzahlStationenCheckAktiv[wpAutomatikkreis]    := 0;
  ailAnzahlFWStationenCheckAktiv[wpAutomatikkreis]  := 0;

  // SHUTTLE
  FOR wlIndex :=   cERSTES_SHUTTLE TO cLETZTES_SHUTTLE DO
    IF StationInAutomatikkreis(starrShuttleBasisParameter[wlIndex].stMKs.eaAutomatikkreis, wpAutomatikkreis) THEN
      starrShuttleBasisParameter[wlIndex].bCheck := FALSE;
      starrShuttleBasisParameter[wlIndex].bCheckMitVorgaenger[cWAND_1] := FALSE;
      starrShuttleBasisParameter[wlIndex].bCheckMitNachfolger[cWAND_1] := FALSE;
    END_IF
  END_FOR

  // STATION
  FOR wlIndex :=   cERSTE_STATION TO cLETZTE_STATION DO
    IF StationInAutomatikkreis(starrStationBasisParameter[wlIndex].stMKs.eaAutomatikkreis, wpAutomatikkreis) THEN
      starrStationBasisParameter[wlIndex].bCheck := FALSE;
      starrStationBasisParameter[wlIndex].bCheckMitVorgaenger[cWAND_1] := FALSE;
      starrStationBasisParameter[wlIndex].bCheckMitNachfolger[cWAND_1] := FALSE;
    END_IF
  END_FOR

  // FW
  FOR wlIndex :=   cERSTE_FAECHERWAGENSTATIONS_NR TO cLETZTE_FAECHERWAGENSTATIONS_NR DO
    IF StationInAutomatikkreis(starrFaecherwagenBasisParameter[wlIndex].stMKs.eaAutomatikkreis, wpAutomatikkreis) THEN
      starrFaecherwagenBasisParameter[wlIndex].bCheck := FALSE;
    END_IF
  END_FOR

  atonlCheckWarteAufMMIDaten[wpAutomatikkreis]( IN :=  FALSE );

  asteplCheck[wpAutomatikkreis, wpZyklus] := STEP_0_E;

END_IF
END_METHOD

(* ---- Vorsteuerung.act.st ---- *)
(* METADATA
{
	"v3Meta": {
		"objectGuid": "2a926ca9-66ff-460d-90cd-a4c06345d8ed"
	}
}
*)
ACTION Vorsteuerung
FOR wlIndexAutomatikkreis := cERSTER_AUTOMATIKKREIS TO cLETZTER_AUTOMATIKKREIS DO

  // Systemcheck aktiv, Zyklen aufteilen
  IF abpCheck[wlIndexAutomatikkreis] THEN

    // Systemcheck starten
    IF NOT ablCheck[wlIndexAutomatikkreis, wlAktiverZyklus] THEN
      ablCheck[wlIndexAutomatikkreis, wlAktiverZyklus] := TRUE;
    END_IF
    // Systemcheck Fehler
    IF ablCheck[wlIndexAutomatikkreis, wlAktiverZyklus] AND abpFehler[wlIndexAutomatikkreis] THEN
      wSps2MmiCheckArea := wlIndexAutomatikkreis;
      wSps2MmiCheckSuccessful := 0;
      MsgToMmi(auftragsnr_w := SB0_SPS_SYSTEMCHECKFINISHED );
      ablCheck[wlIndexAutomatikkreis, wlAktiverZyklus] := FALSE;
      abpCheck[wlIndexAutomatikkreis] := FALSE;
    END_IF
    // Systemcheck abgeschlossen
    IF ablCheck[wlIndexAutomatikkreis, wlAktiverZyklus] AND NOT abpFehler[wlIndexAutomatikkreis] AND ablCheckDone[wlIndexAutomatikkreis, wlAktiverZyklus] THEN
      IF wlAktiverZyklus >= wgAnzahlSystemcheckZyklen THEN
        wSps2MmiCheckArea := wlIndexAutomatikkreis;
        wSps2MmiCheckSuccessful := 1;
        MsgToMmi(auftragsnr_w := SB0_SPS_SYSTEMCHECKFINISHED );
        ablCheck[wlIndexAutomatikkreis, wlAktiverZyklus] := FALSE;
        abpCheck[wlIndexAutomatikkreis] := FALSE;
      ELSE
        // Nächsten Zyklus starten
        ablCheck[wlIndexAutomatikkreis, wlAktiverZyklus] := FALSE;
        wlAktiverZyklus := wlAktiverZyklus + 1;
      END_IF
    END_IF

  // Systemcheck nicht aktiv, alles resetten
  ELSE
    wlAktiverZyklus := 1;
    FOR wlIndexSystemcheckZyklus := 1 TO wgAnzahlSystemcheckZyklen DO
      ablCheck[wlIndexAutomatikkreis, wlIndexSystemcheckZyklus] := FALSE;
    END_FOR
  END_IF

END_FOR
END_ACTION
